PROGRAM main
  VAR
    SCADA_DOOR_OPEN_CMD AT %QX0.0 : BOOL;
    SCADA_DOOR_CLOSE_CMD AT %QX0.1 : BOOL;
    PUB_REMOTE_OPEN_NO_CARD AT %QX0.2 : BOOL;
    PUB_IR_DETECTED AT %QX0.3 : BOOL;
    PUB_DOOR_POSITION AT %QX0.4 : BOOL;
    PUB_ACCESS_GRANTED AT %QX0.5 : BOOL;
    PUB_HEARTBEAT AT %QW0 : UINT;
    PUB_RECONNECT_COUNT AT %QW1 : UINT;
    DOOR_OPEN_CMD AT %QX100.0 : BOOL;
    DOOR_CLOSE_CMD AT %QX100.1 : BOOL;
    IR_DETECTED AT %IX100.0 : BOOL;
    DOOR_POSITION AT %IX100.1 : BOOL;
    ACCESS_GRANTED AT %IX100.2 : BOOL;
    HEARTBEAT AT %IW100 : UINT;
    RECONNECT_COUNT AT %IW101 : UINT;
  END_VAR

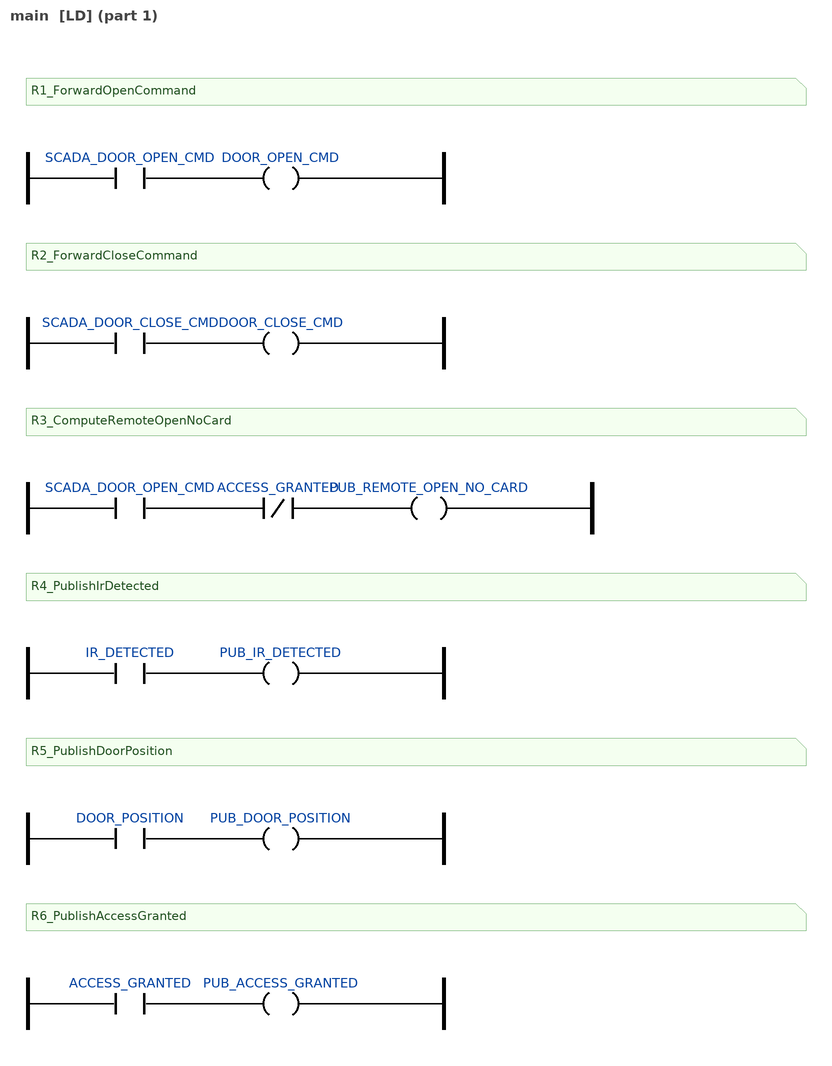
(* LD diagram, written out as Structured Text *)
(* R1_ForwardOpenCommand *)
DOOR_OPEN_CMD := SCADA_DOOR_OPEN_CMD;
(* R2_ForwardCloseCommand *)
DOOR_CLOSE_CMD := SCADA_DOOR_CLOSE_CMD;
(* R3_ComputeRemoteOpenNoCard *)
PUB_REMOTE_OPEN_NO_CARD := SCADA_DOOR_OPEN_CMD AND NOT ACCESS_GRANTED;
(* R4_PublishIrDetected *)
PUB_IR_DETECTED := IR_DETECTED;
(* R5_PublishDoorPosition *)
PUB_DOOR_POSITION := DOOR_POSITION;
(* R6_PublishAccessGranted *)
PUB_ACCESS_GRANTED := ACCESS_GRANTED;
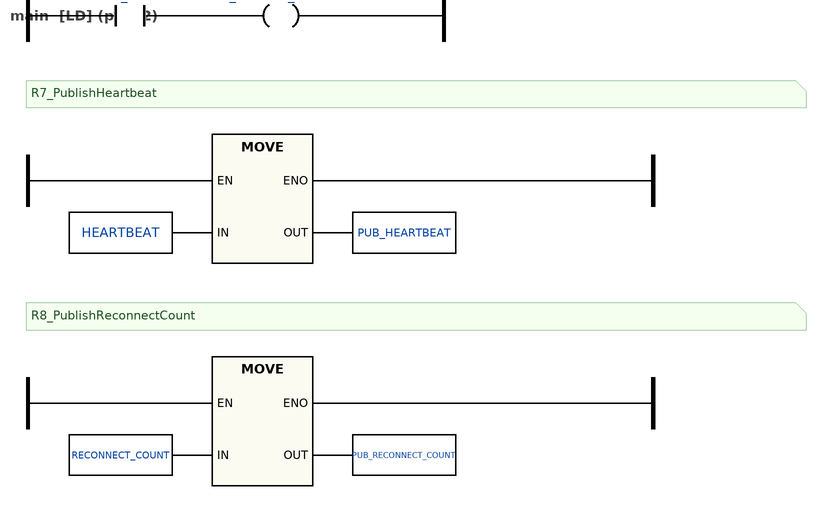
(* R7_PublishHeartbeat *)
PUB_HEARTBEAT := HEARTBEAT;
(* R8_PublishReconnectCount *)
PUB_RECONNECT_COUNT := RECONNECT_COUNT;
END_PROGRAM
